// TIA Portal V20 export
// export: Created 2026-10-12T16:46:20.9204831Z, ExportSetting WithDefaults, DisplayName Totally Integrated Automation Portal, DisplayVersion V20 Update 6, DisplayName TIA Portal Openness, DisplayVersion V20 Update 6, DisplayName TIA Portal Version Control Interface, DisplayVersion V20 Update 6, DisplayName SINAMICS Startdrive Advanced, DisplayVersion V20 SP1 Update 2, DisplayName SINAMICS Startdrive G110M, G120, G120C, G120D, G120P, G115D, DisplayVersion V20 SP1 Update 2, DisplayName SINAMICS Startdrive G130, G150, S120, S150, SINAMICS MV, G220, S200, S210, DisplayVersion V20 SP1 Update 2, DisplayName STEP 7 Professional, DisplayVersion V20 Update 6, DisplayName STEP 7 Safety, DisplayVersion V20 Update 2, DisplayName WinCC Basic/Comfort/Advanced, DisplayVersion V20 Update 6, DisplayName WinCC Professional, DisplayVersion V20 Update 6, DisplayName WinCC Unified, DisplayVersion V20 Update 6
FUNCTION_BLOCK "FB_Heizungssteuerung"   // FB11, SCL
{ S7_Optimized_Access := 'TRUE' }
VERSION : 0.1
// stored: AutoNumber true, IsIECCheckEnabled false, IsRetainMemResEnabled false, MemoryReserve 100, SetENOAutomatically false, UDAEnableTagReadback false
   VAR
      Regler_Bad_7 { S7_SetPoint := 'True'} : "FB_Heizungsregelung";
      Regler_Bad_8 { S7_SetPoint := 'True'} : "FB_Heizungsregelung";
      Regler_Bad_12 { S7_SetPoint := 'True'} : "FB_Heizungsregelung";
      Regler_Bad_25_H1 { S7_SetPoint := 'True'} : "FB_Heizungsregelung";
      Regler_Bad_25_H2 { S7_SetPoint := 'True'} : "FB_Heizungsregelung";
      Regler_Bad_36 { S7_SetPoint := 'True'} : "FB_Heizungsregelung";
      Regler_Bad_40 { S7_SetPoint := 'True'} : "FB_Heizungsregelung";
      Regler_Bad_46 { S7_SetPoint := 'True'} : "FB_Heizungsregelung";
   END_VAR
   VAR_TEMP
      sf : Bool;
   END_VAR
BEGIN

       #sf:="DB_Bad_Konfig".Bad_Konfig[7].IO_Ein.FI_Schutz_OK AND "DB_Bad_Konfig".Bad_Konfig[7].IO_Ein.Kein_Uebertemp AND("DB_Bad_Konfig".Bad_Konfig[7].IO_Ein.Niveau_OK OR NOT "DB_Bad_Konfig".Bad_Konfig[7].Ausstattung.HatNiveau);
       #Regler_Bad_7(Soll:="DB_Bad_Konfig".Bad_Konfig[7].Heizung_1_Soll,Ist:="DB_Bad_Konfig".Bad_Konfig[7].Heizung_1_Ist,Freigabe:=#sf);
       "DB_Bad_Konfig".Bad_Konfig[7].IO_Aus.Heizung_1_Regelung:=#Regler_Bad_7.Schuetz;
       "DB_Bad_Konfig".Bad_Konfig[7].IO_Aus.Heizung_1_Sicherheit:=#sf AND("DB_Bad_Konfig".Bad_Konfig[7].Heizung_1_Soll>0.0);
       #sf:="DB_Bad_Konfig".Bad_Konfig[8].IO_Ein.FI_Schutz_OK AND "DB_Bad_Konfig".Bad_Konfig[8].IO_Ein.Kein_Uebertemp AND("DB_Bad_Konfig".Bad_Konfig[8].IO_Ein.Niveau_OK OR NOT "DB_Bad_Konfig".Bad_Konfig[8].Ausstattung.HatNiveau);
       #Regler_Bad_8(Soll:="DB_Bad_Konfig".Bad_Konfig[8].Heizung_1_Soll,Ist:="DB_Bad_Konfig".Bad_Konfig[8].Heizung_1_Ist,Freigabe:=#sf);
       "DB_Bad_Konfig".Bad_Konfig[8].IO_Aus.Heizung_1_Regelung:=#Regler_Bad_8.Schuetz;
       "DB_Bad_Konfig".Bad_Konfig[8].IO_Aus.Heizung_1_Sicherheit:=#sf AND("DB_Bad_Konfig".Bad_Konfig[8].Heizung_1_Soll>0.0);
       #sf:="DB_Bad_Konfig".Bad_Konfig[12].IO_Ein.FI_Schutz_OK AND "DB_Bad_Konfig".Bad_Konfig[12].IO_Ein.Kein_Uebertemp AND("DB_Bad_Konfig".Bad_Konfig[12].IO_Ein.Niveau_OK OR NOT "DB_Bad_Konfig".Bad_Konfig[12].Ausstattung.HatNiveau);
       #Regler_Bad_12(Soll:="DB_Bad_Konfig".Bad_Konfig[12].Heizung_1_Soll,Ist:="DB_Bad_Konfig".Bad_Konfig[12].Heizung_1_Ist,Freigabe:=#sf);
       "DB_Bad_Konfig".Bad_Konfig[12].IO_Aus.Heizung_1_Regelung:=#Regler_Bad_12.Schuetz;
       "DB_Bad_Konfig".Bad_Konfig[12].IO_Aus.Heizung_1_Sicherheit:=#sf AND("DB_Bad_Konfig".Bad_Konfig[12].Heizung_1_Soll>0.0);
       #sf:="DB_Bad_Konfig".Bad_Konfig[25].IO_Ein.FI_Schutz_OK AND "DB_Bad_Konfig".Bad_Konfig[25].IO_Ein.Kein_Uebertemp AND("DB_Bad_Konfig".Bad_Konfig[25].IO_Ein.Niveau_OK OR NOT "DB_Bad_Konfig".Bad_Konfig[25].Ausstattung.HatNiveau);
       #Regler_Bad_25_H1(Soll:="DB_Bad_Konfig".Bad_Konfig[25].Heizung_1_Soll,Ist:="DB_Bad_Konfig".Bad_Konfig[25].Heizung_1_Ist,Freigabe:=#sf);
       "DB_Bad_Konfig".Bad_Konfig[25].IO_Aus.Heizung_1_Regelung:=#Regler_Bad_25_H1.Schuetz;
       #Regler_Bad_25_H2(Soll:="DB_Bad_Konfig".Bad_Konfig[25].Heizung_2_Soll,Ist:="DB_Bad_Konfig".Bad_Konfig[25].Heizung_2_Ist,Freigabe:=#sf);
       "DB_Bad_Konfig".Bad_Konfig[25].IO_Aus.Heizung_2_Regelung:=#Regler_Bad_25_H2.Schuetz;
       "DB_Bad_Konfig".Bad_Konfig[25].IO_Aus.Heizung_1_Sicherheit:=#sf AND(("DB_Bad_Konfig".Bad_Konfig[25].Heizung_1_Soll>0.0)OR("DB_Bad_Konfig".Bad_Konfig[25].Heizung_2_Soll>0.0));
       "DB_Bad_Konfig".Bad_Konfig[25].IO_Aus.Heizung_2_Sicherheit:="DB_Bad_Konfig".Bad_Konfig[25].IO_Aus.Heizung_1_Sicherheit;
       #sf:="DB_Bad_Konfig".Bad_Konfig[36].IO_Ein.FI_Schutz_OK AND "DB_Bad_Konfig".Bad_Konfig[36].IO_Ein.Kein_Uebertemp AND("DB_Bad_Konfig".Bad_Konfig[36].IO_Ein.Niveau_OK OR NOT "DB_Bad_Konfig".Bad_Konfig[36].Ausstattung.HatNiveau);
       #Regler_Bad_36(Soll:="DB_Bad_Konfig".Bad_Konfig[36].Heizung_1_Soll,Ist:="DB_Bad_Konfig".Bad_Konfig[36].Heizung_1_Ist,Freigabe:=#sf);
       "DB_Bad_Konfig".Bad_Konfig[36].IO_Aus.Heizung_1_Regelung:=#Regler_Bad_36.Schuetz;
       "DB_Bad_Konfig".Bad_Konfig[36].IO_Aus.Heizung_1_Sicherheit:=#sf AND("DB_Bad_Konfig".Bad_Konfig[36].Heizung_1_Soll>0.0);
       #sf:="DB_Bad_Konfig".Bad_Konfig[40].IO_Ein.FI_Schutz_OK AND "DB_Bad_Konfig".Bad_Konfig[40].IO_Ein.Kein_Uebertemp AND("DB_Bad_Konfig".Bad_Konfig[40].IO_Ein.Niveau_OK OR NOT "DB_Bad_Konfig".Bad_Konfig[40].Ausstattung.HatNiveau);
       #Regler_Bad_40(Soll:="DB_Bad_Konfig".Bad_Konfig[40].Heizung_1_Soll,Ist:="DB_Bad_Konfig".Bad_Konfig[40].Heizung_1_Ist,Freigabe:=#sf);
       "DB_Bad_Konfig".Bad_Konfig[40].IO_Aus.Heizung_1_Regelung:=#Regler_Bad_40.Schuetz;
       "DB_Bad_Konfig".Bad_Konfig[40].IO_Aus.Heizung_1_Sicherheit:=#sf AND("DB_Bad_Konfig".Bad_Konfig[40].Heizung_1_Soll>0.0);
       #sf:="DB_Bad_Konfig".Bad_Konfig[46].IO_Ein.FI_Schutz_OK AND "DB_Bad_Konfig".Bad_Konfig[46].IO_Ein.Kein_Uebertemp AND("DB_Bad_Konfig".Bad_Konfig[46].IO_Ein.Niveau_OK OR NOT "DB_Bad_Konfig".Bad_Konfig[46].Ausstattung.HatNiveau);
       #Regler_Bad_46(Soll:="DB_Bad_Konfig".Bad_Konfig[46].Heizung_1_Soll,Ist:="DB_Bad_Konfig".Bad_Konfig[46].Heizung_1_Ist,Freigabe:=#sf);
       "DB_Bad_Konfig".Bad_Konfig[46].IO_Aus.Heizung_1_Regelung:=#Regler_Bad_46.Schuetz;
       "DB_Bad_Konfig".Bad_Konfig[46].IO_Aus.Heizung_1_Sicherheit:=#sf AND("DB_Bad_Konfig".Bad_Konfig[46].Heizung_1_Soll>0.0);
END_FUNCTION_BLOCK
